PROGRAM main
  VAR
    stop : BOOL;
    start : BOOL;
    motor_run : BOOL;
    star : BOOL;
    TON0 : TON;
    delta : BOOL;
    TON1 : TON;
    overload : BOOL;
    red_lamp : BOOL;
  END_VAR

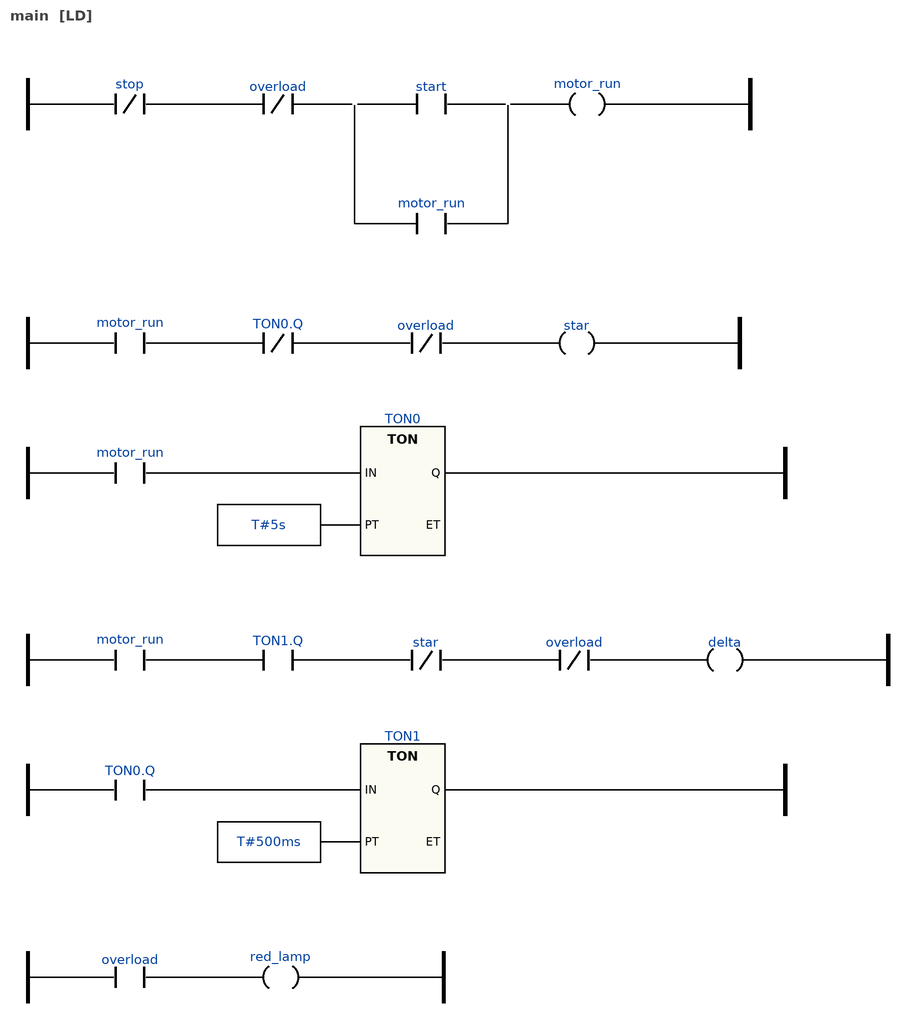
(* LD diagram, written out as Structured Text *)
motor_run := NOT stop AND NOT overload AND (start OR motor_run);
star := motor_run AND NOT TON0.Q AND NOT overload;
delta := motor_run AND TON1.Q AND NOT star AND NOT overload;
red_lamp := overload;
TON0(IN := motor_run, PT := T#5s);
TON1(IN := TON0.Q, PT := T#500ms);
END_PROGRAM
